Fanuc KAREL source: ko00049.KL

-- PROVISIONAL review KL for V770-1; original PC SHA256 1000af24aa73f09ac404206c1b0f1dcc664484904d7ec018f2703fe0f2a45d8c
-- Incomplete behavior may be omitted. Consult companion uncertainty JSON. Do not deploy.
PROGRAM KO00049
%NOLOCKGROUP
BEGIN
  -- UNRESOLVED_PC offsets 5-12; opcodes 9D,23
  -- UNRESOLVED_PC offsets 17-66; opcodes 27,27,49,7E,AD,22,1C,22,31,7E,4A
  -- UNRESOLVED_PC offsets 71-75; opcodes 7F
END KO00049
